(* IEC 61131-3 sources: SemantiST/benchmarks/oscat/targets/oscat_network_ip4_check, 2 files *)

(* ---- normalized.st ---- *)
FUNCTION IP4_CHECK : BOOL
VAR_INPUT
	NIP : DWORD;
	LIP : DWORD;
	SM : DWORD;
END_VAR

(*
version 1.0	4. mar 2008
programmer 	hugo
tested by		oscat

IP4_CHECK testet ob eine Network IP und Local_IP im selben Subnet sind.

*)

IP4_CHECK := (NIP AND sm) = (LIP AND SM);

(* revision history
hm		4. mar 2008	rev 1.0
	original version

*)
END_FUNCTION

(* ---- target.st ---- *)
FUNCTION IP4_CHECK : BOOL
VAR_INPUT
	NIP : DWORD;
	LIP : DWORD;
	SM : DWORD;
END_VAR

(*
version 1.0	4. mar 2008
programmer 	hugo
tested by		oscat

IP4_CHECK testet ob eine Network IP und Local_IP im selben Subnet sind.

*)

IP4_CHECK := (NIP AND sm) = (LIP AND SM);

(* revision history
hm		4. mar 2008	rev 1.0
	original version

*)
END_FUNCTION
